Staubli VAL3: stop.pgx

program stop()
  local num l_nI
begin
  //应用停止时调用：清掉 9 个功能按钮的选中态，避免下次启动带着上次的状态
  for l_nI=0 to 8
    bFunc[l_nI]=false
    sFuncBg[l_nI]="#DCDCDC"
  endFor
end
